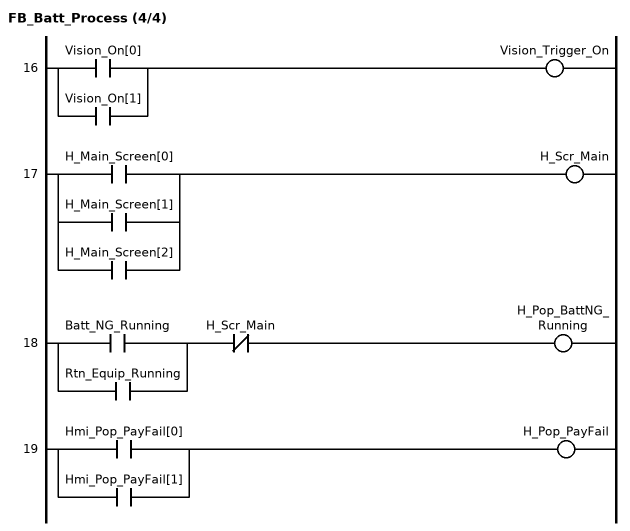
(* [picture p24: FB_Batt_Process, rungs 16-19] *)
(* Rung 16 *)
Vision_Trigger_On := Vision_On[0] OR Vision_On[1];
(* Rung 17 *)
H_Scr_Main := H_Main_Screen[0] OR H_Main_Screen[1] OR H_Main_Screen[2];
(* Rung 18 *)
H_Pop_BattNG_Running := (Batt_NG_Running OR Rtn_Equip_Running) AND NOT H_Scr_Main;
(* Rung 19 *)
H_Pop_PayFail := Hmi_Pop_PayFail[0] OR Hmi_Pop_PayFail[1];
END_FUNCTION_BLOCK

FUNCTION_BLOCK Connect
VAR
    nStep : INT := 0;
    exAccept : BOOL;
    exRcv : BOOL;
    exSend : BOOL;
    exClose : BOOL;
    TCP_Accept : SktTCPAccept;
    TCP_Recv : SktTCPRcv;
    TCP_Send : SktTCPSend;
    TCP_Close : SktClose;
    Sock : _sSOCKET;
    RxBuf : ARRAY[0..259] OF BYTE;
    TxBuf : ARRAY[0..259] OF BYTE;
    TxSize : UINT;
    FC : BYTE;
    Addr : UINT;
    Qty : UINT;
    i : UINT;
    ExCode : BYTE;
    RetryT : TON;
    HR_SIZE : UINT := 100;
    ErrStep : INT;
END_VAR
VAR_INPUT
    Enable : BOOL;  (* TRUE면 서버 동작 *)
    Port : UINT;  (* 대기할 TCP 포트 번호 (MFC 502 / 아두이노 503) *)
END_VAR
VAR_IN_OUT
    HR : ARRAY[0..99] OF WORD;  (* Modbus 레지스터 0~99번 *)
END_VAR
VAR_OUTPUT
    Connected : BOOL;  (* 클라이언트 접속 중 *)
    ErrorID : WORD;  (* 마지막 에러 코드 *)
    ReqCount : UDINT;  (* 처리한 요청 수 (통신 확인용) *)
END_VAR
CASE nStep OF

    0 : (*정지 상태*)
    Connected := FALSE;
    IF Enable THEN
        nStep := 10;
    END_IF;

    10 : (*클라이언트 접속 대기*)
    exAccept := TRUE;
    IF TCP_Accept.Done THEN
        exAccept := FALSE;
        Sock:=TCP_Accept.Socket;
        Connected := TRUE;
		ErrorID := WORD#16#0;
		ErrStep := 0;
        nStep := 20;
	ELSIF TCP_Accept.Error THEN
		exAccept := FALSE;
		ErrorID := TCP_Accept.ErrorID;
		ErrStep := 10;
		nStep := 90;
    END_IF;

    20 : (*요청 수신*)
    exRcv:=TRUE;
    IF TCP_Recv.Done THEN
        exRcv := FALSE;
        IF TCP_Recv.RcvSize = UINT#0 THEN
            nStep := 80; (*클라이언트에 의한 연결 종료*)
        ELSIF TCP_Recv.RcvSize >= UINT#12 THEN
            nStep := 30; (*정상 수신*)
        END_IF;
    ELSIF TCP_Recv.Error THEN
        exRcv :=FALSE;
        ErrorID := TCP_Recv.ErrorID;
		ErrStep := 20;
        nStep := 80;
    END_IF;

    30 : (*요청 해석 = 응답 작성*)
    FC := RxBuf[7];
    Addr := BYTE_TO_UINT(RxBuf[8]) * UINT#256 + BYTE_TO_UINT(RxBuf[9]);
    Qty := BYTE_TO_UINT(RxBuf[10]) * UINT#256 + BYTE_TO_UINT(RxBuf[11]);
    ExCode := BYTE#16#00;

    FOR i := UINT#0 TO UINT#6 DO
        TxBuf[i] := RxBuf[i];
    END_FOR;
    TxBuf[7] := FC;

    IF FC = BYTE#16#03 THEN (*Holding Register 읽기*)
        IF (Qty < UINT#1) OR (Qty > UINT#125) THEN
            ExCode := BYTE#16#03;
        ELSIF (Addr + Qty) > HR_SIZE THEN
            ExCode := BYTE#16#02;
        ELSE
            TxBuf[8] := UINT_TO_BYTE(Qty * UINT#2);
            FOR i := UINT#0 TO Qty - UINT#1 DO
                TxBuf[UINT#9 + i * UINT#2] := WORD_TO_BYTE(SHR(HR[Addr + i], 8));
                TxBuf[UINT#10 + i * UINT#2] := WORD_TO_BYTE(HR[Addr + i]);
            END_FOR;
            TxSize := UINT#9 + Qty * UINT#2;
        END_IF;
    ELSIF FC = BYTE#16#06 THEN (*Register 작성 - 1개*)
        IF Addr >= HR_SIZE THEN
            ExCode := BYTE#16#02;
        ELSE
            HR[Addr] := UINT_TO_WORD(Qty);
            FOR i := UINT#8 TO UINT#11 DO
                TxBuf[i] := RxBuf[i];
            END_FOR;
            TxSize := UINT#12;
        END_IF;
    ELSIF FC = BYTE#16#10 THEN (*Register 작성 - 복수*)
        IF (Qty < UINT#1) OR (Qty > UINT#123) OR (BYTE_TO_UINT(RxBuf[12]) <> Qty * UINT#2) OR (TCP_Recv.RcvSize < UINT#13 + Qty * UINT#2) THEN
            ExCode := BYTE#16#03;
        ELSIF (Addr + Qty) > HR_SIZE THEN
            ExCode := BYTE#16#02;
        ELSE
            FOR i := UINT#0 TO Qty - UINT#1 DO
                HR[Addr + i] := UINT_TO_WORD(BYTE_TO_UINT(RxBuf[UINT#13 + i * UINT#2]) * UINT#256 + BYTE_TO_UINT(RxBuf[UINT#14 + i * UINT#2]));
            END_FOR;    
            FOR i := UINT#8 TO UINT#11 DO
                TxBuf[i] := RxBuf[i]; (*시작 주소 + 개수*)
            END_FOR;
            TxSize := UINT#12;
        END_IF;
    ELSE
        ExCode := BYTE#16#01; (*지원하지 않는 기능 코드*)
    END_IF;

    IF ExCode <> BYTE#16#00 THEN (*예외 응답*)
        TxBuf[7] := FC OR BYTE#16#80;
        TxBuf[8] := ExCode;
        TxSize := UINT#9;
    END_IF;

    (*바이트 수 - 유닛 ID부터 끝까지*)
    TxBuf[4] := BYTE#16#00;
    TxBuf[5] := UINT_TO_BYTE(TxSize - UINT#6);
    nStep := 40;

    40 : (*응답 송신*)
    exSend := TRUE;
    IF TCP_Send.Done THEN
        exSend := FALSE;
        ReqCount := ReqCount + UDINT#1;
        nStep := 20; (*다음 요청 대기*)
    ELSIF TCP_Send.Error THEN
        exSend :=FALSE;
        ErrorID := TCP_Send.ErrorID;
        nStep := 80;
    END_IF;

    80 : (*소켓 CLOSE*)
    exClose := TRUE;
    Connected := FALSE;
    IF TCP_Close.Done THEN
        exClose := FALSE;
        nStep := 90;
	ELSIF TCP_Close.Error THEN
		exClose := FALSE;
		IF ErrorID = WORD#16#0 THEN
			ErrorID := TCP_Close.ErrorID;
			ErrStep := 80;
		END_IF;
		nStep := 90;
    END_IF;

    90 : (*1초 후 재접속 대기*)
    IF RetryT.Q THEN
        nStep := 0;
    END_IF;

END_CASE;

(*명령 호출*)
TCP_Accept(Execute := exAccept, SrcTcpPort := Port, TimeOut := UINT#0);
TCP_Recv(Execute := exRcv, Socket := Sock, TimeOut := UINT#50, Size := UINT#260, RcvDat := RxBuf[0]);
TCP_Send(Execute := exSend, Socket := Sock, SendDat := TxBuf[0], Size := TxSize);
TCP_Close(Execute := exClose, Socket := Sock);
RetryT(In := (nStep = 90), PT := T#1s);
END_FUNCTION_BLOCK

# Device HMI_NA5_0 (NA): not converted